// TIA Portal project "DistributoreCaffè" (V19)

(* hardware
DEVICE "S7-1200 station_1"  S7-1200 Station
   slot 0: "Telaio di montaggio_0"  S7-1200 Rack  Rack  V1.0
   slot 1: "PLC"  CPU 1212C DC/DC/Rly  6ES7 212-1HE40-0XB0  V4.6
DEVICE "HMI"  KTP900 Basic PN
   slot 0: "HMI_1"  KTP900 Basic PN  6AV2 123-2JB03-0AX0  17.0.0.0
   slot 1: "HMI_RT_1"  KTP900 Basic PN  6AV2 123-2JB03-0AX0  17.0.0.0
   slot 5: "HMI_1.IE_CP_1"  PROFINET Interface  17.0.0.0
      slot 1: "Interfaccia_1 PROFINET"  PROFINET Interface
         slot 1: "Porta_1"  Port
*)

// ===== PLC "PLC"  CPU 1212C DC/DC/Rly =====

TYPE "CreditoResto"
   STRUCT
      "5Cents" : Real;
      "10Cents" : Real;
      "20Cents" : Real;
      "50Cents" : Real;
      "1Euro" : Real;
      "2Euro" : Real;
   END_STRUCT;
END_TYPE

TYPE "RestoUtente"
   STRUCT
      "5Cents" : SInt;
      "10Cents" : SInt;
      "20Cents" : SInt;
      "50Cents" : SInt;
      "1Euro" : SInt;
      "2Euro" : SInt;
   END_STRUCT;
END_TYPE

TYPE "Prezzo"
   STRUCT
      Bevanda : String;
      Prezzo : Real;
   END_STRUCT;
END_TYPE

DATA_BLOCK "HMI"   // DB1
{ S7_Optimized_Access := 'TRUE' }
VERSION : 0.1
   VAR
      I5cents : Bool;
      I10Cents : Bool;
      I20Cents : Bool;
      I50Cents : Bool;
      I1Euro : Bool;
      I2Euro : Bool;
   END_VAR
   VAR RETAIN
      Resto : "RestoUtente";
   END_VAR
   VAR
      ValvolaBicchiere : Bool;
      ValvolaPaletta : Bool;
      ValvolaCaffè : Bool;
      ValvolaLatte : Bool;
      ValvolaGrappa : Bool;
      ValvolaZucchero : Bool;
      PrelievoProdotto : Bool;
   END_VAR
   VAR RETAIN
      ProdottoPronto : Bool;
   END_VAR
   VAR
      Corto : Bool;
      CortoMacchiato : Bool;
      CortoCorretto : Bool;
      CortoMacchiatoCorretto : Bool;
      Lungo : Bool;
      LungoMacchiato : Bool;
      LungoCorretto : Bool;
      LungoMacchiatoCorretto : Bool;
      ConfermaOrdine : Bool;
      BicchieriScarico : Bool;
      PaletteScarico : Bool;
      CaffèScarico : Bool;
      LatteScarico : Bool;
      GrappaScarico : Bool;
      ZuccheroScarico : Bool;
      Bicchieri : Int;
      Palette : Int;
      Caffè : SInt;
      Latte : SInt;
      Grappa : SInt;
      Zucchero : SInt;
   END_VAR
   VAR RETAIN
      Credito : Real;
      Introiti : Real;
   END_VAR
   VAR
      PrelievoIntroiti : Bool;
      CreditoInsufficiente : Bool;
      QuantitàZuccheroSelezionata : SInt;
      RiduzioneZucchero : Bool;
      IncrementoZucchero : Bool;
      ProdottoInPreparazione : Bool;
   END_VAR
BEGIN
END_DATA_BLOCK

DATA_BLOCK "Sistema"   // DB2
{ S7_Optimized_Access := 'TRUE' }
VERSION : 0.1
   VAR RETAIN
      CreditoResto : "CreditoResto";
   END_VAR
   VAR
      PConfermaOrdine : Bool;
      BloccoInterfacciaUtente : Bool;
      NPrelievoProdotto : Bool;
      BevandaSelezionata : SInt;
      PCorto : Bool;
      PCortoMacchiato : Bool;
      PCortoCorretto : Bool;
      PCortoMacchiatoCorretto : Bool;
      PLungo : Bool;
      PLungoMacchiato : Bool;
      PLungoCorretto : Bool;
      PLungoMacchiatoCorretto : Bool;
      PPiùZucchero : Bool;
      PMenoZucchero : Bool;
   END_VAR
   VAR RETAIN
      Prezzi : Array[1..8] of "Prezzo";
   END_VAR
   VAR
      PBloccoInterfacciaUtente : Bool;
      NPrelievoProdotto2 : Bool;
      NPrelievoIntroiti : Bool;
   END_VAR
BEGIN
   CreditoResto."5Cents" := 5.0;
   CreditoResto."10Cents" := 5.0;
   CreditoResto."20Cents" := 5.0;
   CreditoResto."50Cents" := 5.0;
   CreditoResto."1Euro" := 5.0;
   CreditoResto."2Euro" := 5.0;
   Prezzi[1].Bevanda := 'Corto';
   Prezzi[1].Prezzo := 0.3;
   Prezzi[2].Bevanda := 'CortoMacchiato';
   Prezzi[2].Prezzo := 0.4;
   Prezzi[3].Bevanda := 'CortoCorretto';
   Prezzi[3].Prezzo := 0.4;
   Prezzi[4].Bevanda := 'CortoMacchiatoCorretto';
   Prezzi[4].Prezzo := 0.5;
   Prezzi[5].Bevanda := 'Lungo';
   Prezzi[5].Prezzo := 0.6;
   Prezzi[6].Bevanda := 'LungoMacchiato';
   Prezzi[6].Prezzo := 0.7;
   Prezzi[7].Bevanda := 'LungoCorretto';
   Prezzi[7].Prezzo := 0.7;
   Prezzi[8].Bevanda := 'LungoMacchiatoCorretto';
   Prezzi[8].Prezzo := 0.8;
END_DATA_BLOCK

DATA_BLOCK "AggiornamentoCreditoUtente_DB"   // DB3
{ S7_Optimized_Access := 'TRUE' }
VERSION : 0.1
// stored: InstanceOfName AggiornamentoCreditoUtenteCreditoDistributore
"AggiornamentoCreditoUtenteCreditoDistributore"
BEGIN
END_DATA_BLOCK

DATA_BLOCK "PreparazioneBevanda_DB"   // DB4
{ S7_Optimized_Access := 'TRUE' }
VERSION : 0.1
// stored: InstanceOfName PreparazioneBevanda
"PreparazioneBevanda"
BEGIN
END_DATA_BLOCK

DATA_BLOCK "AggiornamentoRestoUtenteCreditoUtenteCreditoDistributore_DB"   // DB5
{ S7_Optimized_Access := 'TRUE' }
VERSION : 0.1
// stored: InstanceOfName AggiornamentoRestoUtenteCreditoUtenteCreditoDistributore
"AggiornamentoRestoUtenteCreditoUtenteCreditoDistributore"
BEGIN
END_DATA_BLOCK

FUNCTION_BLOCK "AggiornamentoCreditoUtenteCreditoDistributore"   // FB1, LAD
{ S7_Optimized_Access := 'TRUE' }
VERSION : 0.1
   VAR_INPUT
      "5Cents" : Bool;
      "10Cents" : Bool;
      "20Cents" : Bool;
      "50Cents" : Bool;
      "1Euro" : Bool;
      "2Euro" : Bool;
   END_VAR
   VAR_IN_OUT
      CreditoDistributore : "CreditoResto";
      CreditoUtente : Real;
   END_VAR
   VAR
      PI5Cents : Bool;
      PI10Cents : Bool;
      PI20Cents : Bool;
      PI50Cents : Bool;
      PI1Euro : Bool;
      PI2Euro : Bool;
   END_VAR
   VAR_TEMP   // added for the SCL form of the ladder/FBD networks
      _w1 : Bool;
      _w2 : Bool;
      _w3 : Bool;
      _w4 : Bool;
      _w5 : Bool;
      _w6 : Bool;
   END_VAR
BEGIN

REGION Network 1
   // Attenzione: i valori Real non sempre vengono salvati a cifra tonda
   // (Es: 0.2999999999.. oppure 0.31111111.. invece di 0.3)
   // Arrotondare dopo ogni operazione matematica che li implica
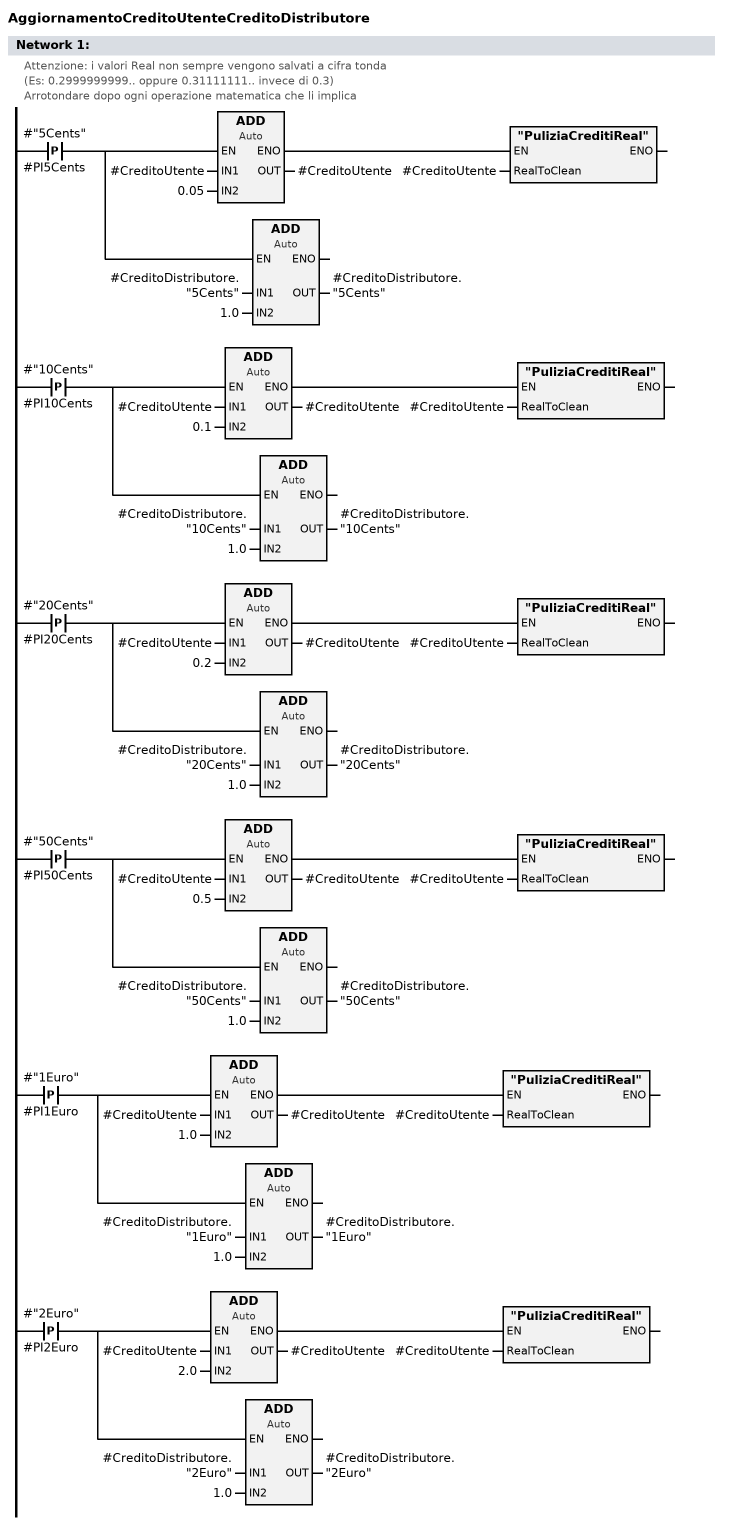
   RUNG wire#powerrail
      P_Contact(operand := #"5Cents", bit := #PI5Cents)
      wire#w1
      Add(in1 := #CreditoUtente, in2 := 0.05, out => #CreditoUtente)
      "PuliziaCreditiReal"(RealToClean := #CreditoUtente)
   END_RUNG
   RUNG wire#w1
      Add(in1 := #CreditoDistributore."5Cents", in2 := 1.0, out => #CreditoDistributore."5Cents")
   END_RUNG
   RUNG wire#powerrail
      P_Contact(operand := #"10Cents", bit := #PI10Cents)
      wire#w2
      Add(in1 := #CreditoUtente, in2 := 0.1, out => #CreditoUtente)
      "PuliziaCreditiReal"(RealToClean := #CreditoUtente)
   END_RUNG
   RUNG wire#w2
      Add(in1 := #CreditoDistributore."10Cents", in2 := 1.0, out => #CreditoDistributore."10Cents")
   END_RUNG
   RUNG wire#powerrail
      P_Contact(operand := #"20Cents", bit := #PI20Cents)
      wire#w3
      Add(in1 := #CreditoUtente, in2 := 0.2, out => #CreditoUtente)
      "PuliziaCreditiReal"(RealToClean := #CreditoUtente)
   END_RUNG
   RUNG wire#w3
      Add(in1 := #CreditoDistributore."20Cents", in2 := 1.0, out => #CreditoDistributore."20Cents")
   END_RUNG
   RUNG wire#powerrail
      P_Contact(operand := #"50Cents", bit := #PI50Cents)
      wire#w4
      Add(in1 := #CreditoUtente, in2 := 0.5, out => #CreditoUtente)
      "PuliziaCreditiReal"(RealToClean := #CreditoUtente)
   END_RUNG
   RUNG wire#w4
      Add(in1 := #CreditoDistributore."50Cents", in2 := 1.0, out => #CreditoDistributore."50Cents")
   END_RUNG
   RUNG wire#powerrail
      P_Contact(operand := #"1Euro", bit := #PI1Euro)
      wire#w5
      Add(in1 := #CreditoUtente, in2 := 1.0, out => #CreditoUtente)
      "PuliziaCreditiReal"(RealToClean := #CreditoUtente)
   END_RUNG
   RUNG wire#w5
      Add(in1 := #CreditoDistributore."1Euro", in2 := 1.0, out => #CreditoDistributore."1Euro")
   END_RUNG
   RUNG wire#powerrail
      P_Contact(operand := #"2Euro", bit := #PI2Euro)
      wire#w6
      Add(in1 := #CreditoUtente, in2 := 2.0, out => #CreditoUtente)
      "PuliziaCreditiReal"(RealToClean := #CreditoUtente)
   END_RUNG
   RUNG wire#w6
      Add(in1 := #CreditoDistributore."2Euro", in2 := 1.0, out => #CreditoDistributore."2Euro")
   END_RUNG
   // the same network as SCL:
   #_w1 := #"5Cents" AND NOT #PI5Cents;   // rising edge of #"5Cents"
   #PI5Cents := #"5Cents";
   IF #_w1 THEN
       #CreditoUtente := #CreditoUtente + 0.05;
       "PuliziaCreditiReal"(RealToClean := #CreditoUtente);
       #CreditoDistributore."5Cents" := #CreditoDistributore."5Cents" + 1.0;
   END_IF;
   #_w2 := #"10Cents" AND NOT #PI10Cents;   // rising edge of #"10Cents"
   #PI10Cents := #"10Cents";
   IF #_w2 THEN
       #CreditoUtente := #CreditoUtente + 0.1;
       "PuliziaCreditiReal"(RealToClean := #CreditoUtente);
       #CreditoDistributore."10Cents" := #CreditoDistributore."10Cents" + 1.0;
   END_IF;
   #_w3 := #"20Cents" AND NOT #PI20Cents;   // rising edge of #"20Cents"
   #PI20Cents := #"20Cents";
   IF #_w3 THEN
       #CreditoUtente := #CreditoUtente + 0.2;
       "PuliziaCreditiReal"(RealToClean := #CreditoUtente);
       #CreditoDistributore."20Cents" := #CreditoDistributore."20Cents" + 1.0;
   END_IF;
   #_w4 := #"50Cents" AND NOT #PI50Cents;   // rising edge of #"50Cents"
   #PI50Cents := #"50Cents";
   IF #_w4 THEN
       #CreditoUtente := #CreditoUtente + 0.5;
       "PuliziaCreditiReal"(RealToClean := #CreditoUtente);
       #CreditoDistributore."50Cents" := #CreditoDistributore."50Cents" + 1.0;
   END_IF;
   #_w5 := #"1Euro" AND NOT #PI1Euro;   // rising edge of #"1Euro"
   #PI1Euro := #"1Euro";
   IF #_w5 THEN
       #CreditoUtente := #CreditoUtente + 1.0;
       "PuliziaCreditiReal"(RealToClean := #CreditoUtente);
       #CreditoDistributore."1Euro" := #CreditoDistributore."1Euro" + 1.0;
   END_IF;
   #_w6 := #"2Euro" AND NOT #PI2Euro;   // rising edge of #"2Euro"
   #PI2Euro := #"2Euro";
   IF #_w6 THEN
       #CreditoUtente := #CreditoUtente + 2.0;
       "PuliziaCreditiReal"(RealToClean := #CreditoUtente);
       #CreditoDistributore."2Euro" := #CreditoDistributore."2Euro" + 1.0;
   END_IF;
END_REGION
END_FUNCTION_BLOCK

FUNCTION_BLOCK "PreparazioneBevanda"   // FB2, LAD
{ S7_Optimized_Access := 'TRUE' }
VERSION : 0.1
   VAR_INPUT
      BevandaSelezionata : SInt;
      InnescoProcesso : Bool;
   END_VAR
   VAR
      TPBicchiere : TP_TIME;
      NQTPBicchiere : Bool;
      TPPaletta : TP_TIME;
      NQTPPaletta : Bool;
      TPCaffè : TP_TIME;
      NQTPCaffè : Bool;
      TPLatte : TP_TIME;
      NQTPLatte : Bool;
      TPGrappa : TP_TIME;
      NQTPGrappa : Bool;
      TPzucchero : TP_TIME;
      NQTPZucchero : Bool;
      PInnescoProcesso : Bool;
   END_VAR
   VAR_TEMP
      PTZucchero : Int;
   END_VAR
   VAR_TEMP   // added for the SCL form of the ladder/FBD networks
      _w1 : Bool;
      _w2 : Bool;
      _w3 : Bool;
      _w4 : Bool;
      _w5 : Bool;
      _w6 : Bool;
      _w7 : Bool;
      _w8 : Bool;
      _w9 : Bool;
      _w10 : Bool;
      _w11 : Bool;
      _w12 : Bool;
   END_VAR
BEGIN

REGION Network 1
   // Gestire trigger timer valvole
   // - grappa caso bevanda corretta non macchiata
   // - zucchero caso bevanda zuccherata liscia o macchiata
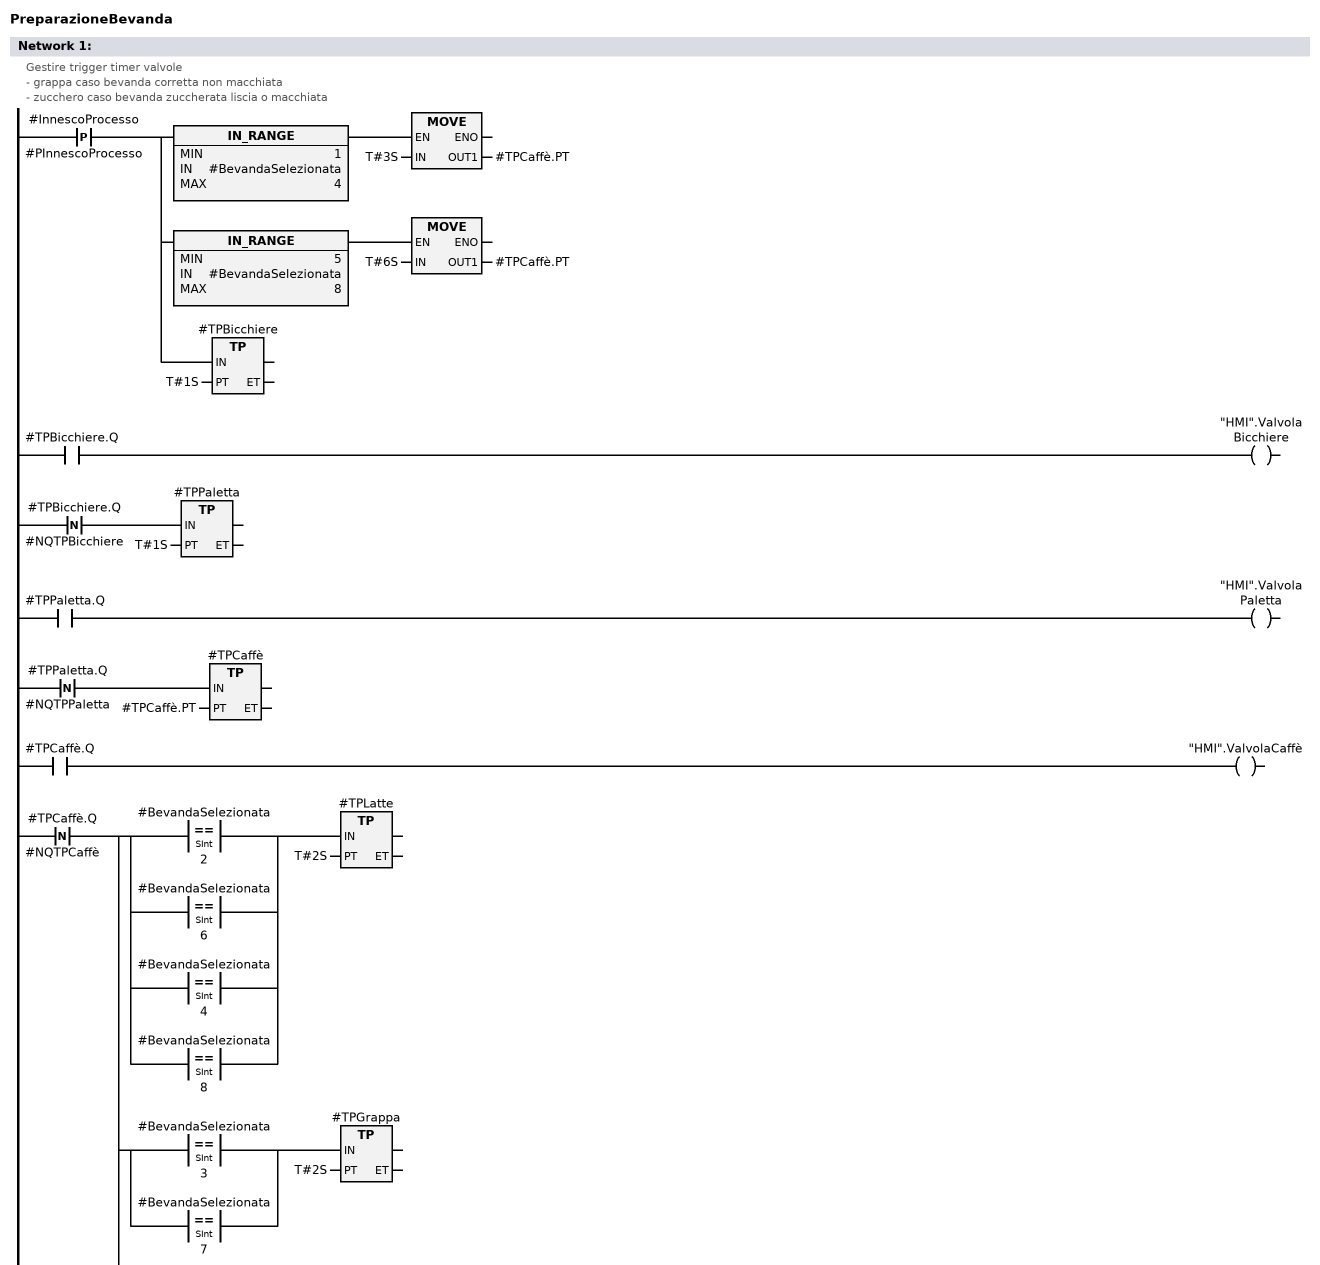
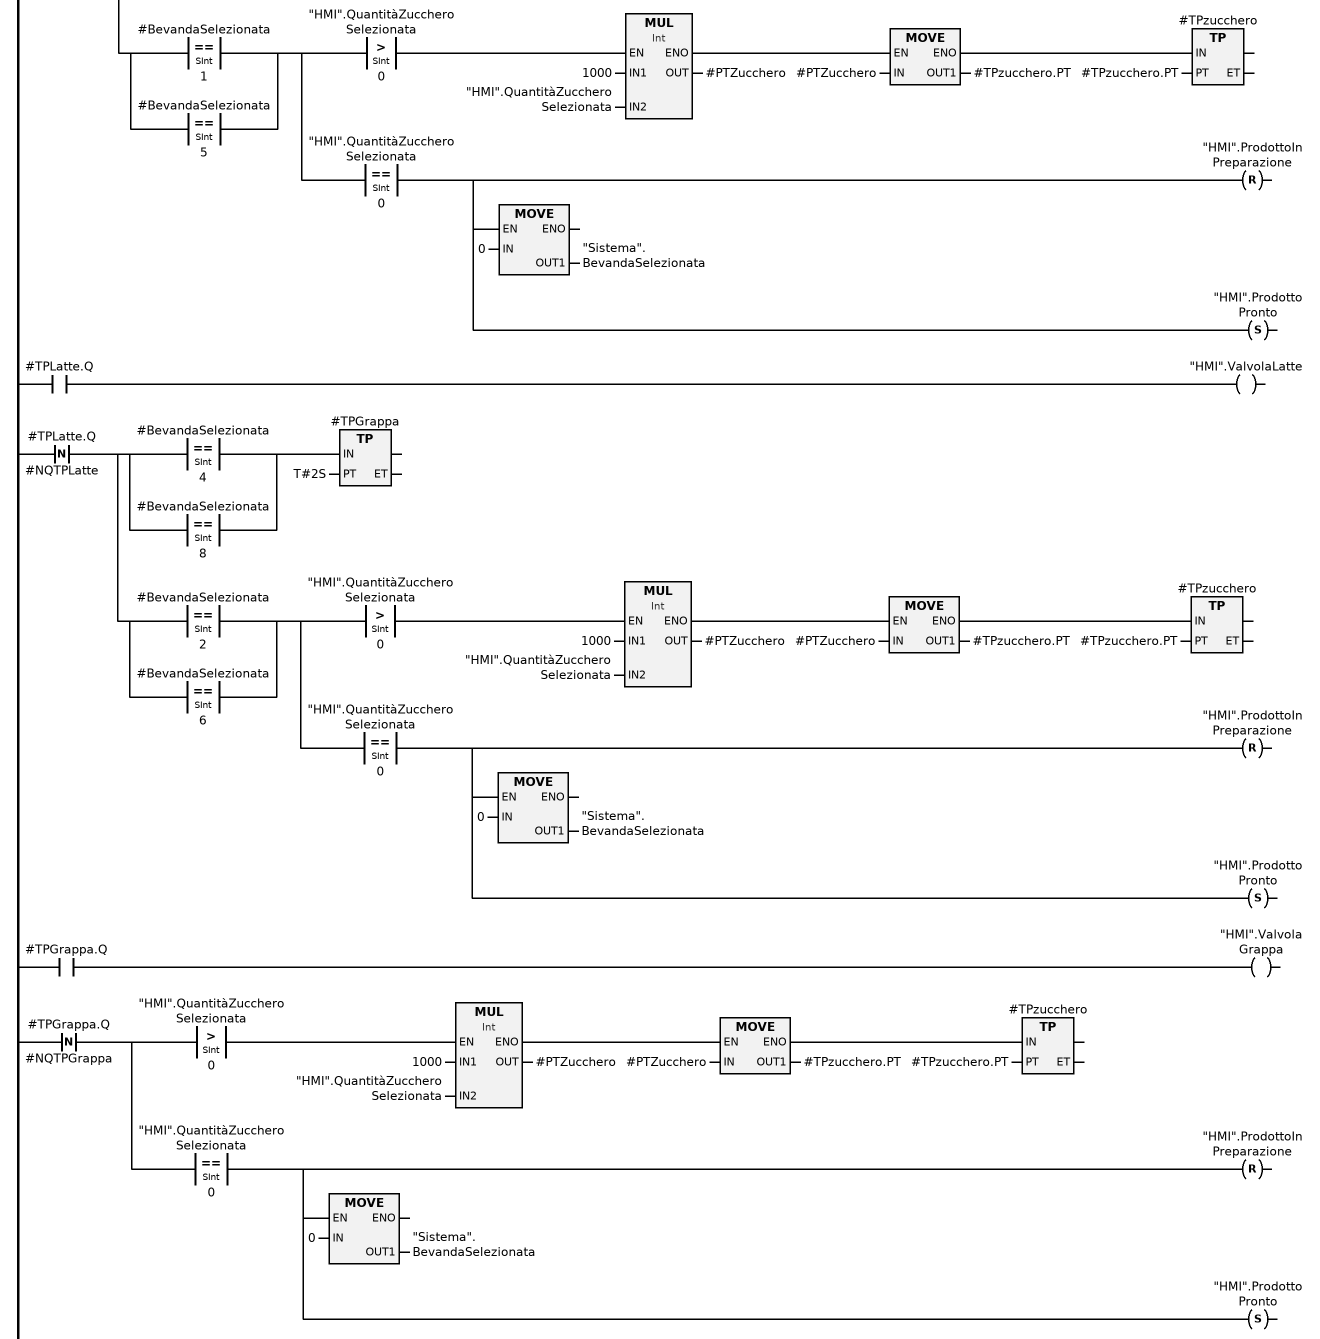
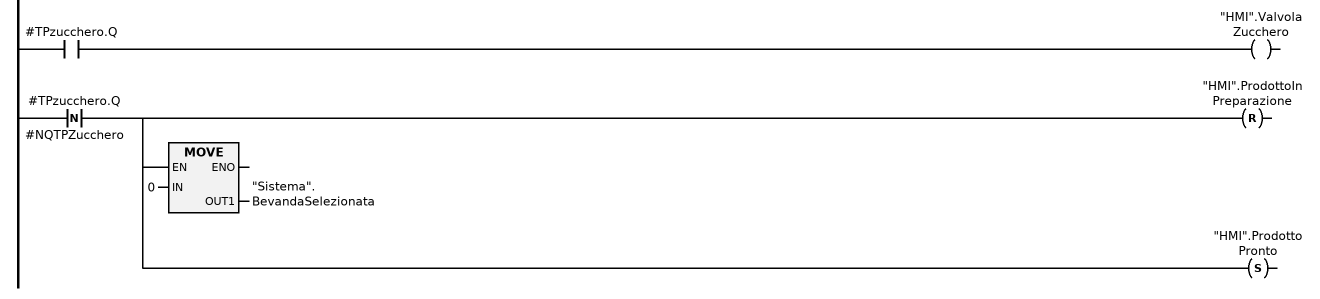
   #_w1 := #InnescoProcesso AND NOT #PInnescoProcesso;   // rising edge of #InnescoProcesso
   #PInnescoProcesso := #InnescoProcesso;
   IF #_w1 AND (1 <= #BevandaSelezionata) AND (#BevandaSelezionata <= 4) THEN #TPCaffè.PT := T#3S; END_IF;
   IF #_w1 AND (5 <= #BevandaSelezionata) AND (#BevandaSelezionata <= 8) THEN #TPCaffè.PT := T#6S; END_IF;
   #TPBicchiere(IN := #_w1, PT := T#1S);   // TP
   "HMI".ValvolaBicchiere := #TPBicchiere.Q;
   #_w2 := NOT #TPBicchiere.Q AND #NQTPBicchiere;   // falling edge of #TPBicchiere.Q
   #NQTPBicchiere := #TPBicchiere.Q;
   #TPPaletta(IN := #_w2, PT := T#1S);   // TP
   "HMI".ValvolaPaletta := #TPPaletta.Q;
   #_w3 := NOT #TPPaletta.Q AND #NQTPPaletta;   // falling edge of #TPPaletta.Q
   #NQTPPaletta := #TPPaletta.Q;
   #TPCaffè(IN := #_w3, PT := #TPCaffè.PT);   // TP
   "HMI".ValvolaCaffè := #TPCaffè.Q;
   #_w4 := NOT #TPCaffè.Q AND #NQTPCaffè;   // falling edge of #TPCaffè.Q
   #NQTPCaffè := #TPCaffè.Q;
   #TPLatte(IN := #_w4 AND ((#BevandaSelezionata = 2) OR (#BevandaSelezionata = 6) OR (#BevandaSelezionata = 4) OR (#BevandaSelezionata = 8)),   // TP
            PT := T#2S);
   #TPGrappa(IN := #_w4 AND ((#BevandaSelezionata = 3) OR (#BevandaSelezionata = 7)), PT := T#2S);   // TP
   #_w5 := #_w4 AND ((#BevandaSelezionata = 1) OR (#BevandaSelezionata = 5));
   #_w6 := #_w5 AND ("HMI".QuantitàZuccheroSelezionata > 0);
   IF #_w6 THEN
       #PTZucchero := 1000 * "HMI".QuantitàZuccheroSelezionata;
       #TPzucchero.PT := #PTZucchero;
   END_IF;
   #TPzucchero(IN := #_w6, PT := #TPzucchero.PT);   // TP
   IF #_w5 AND ("HMI".QuantitàZuccheroSelezionata = 0) THEN
       "HMI".ProdottoInPreparazione := FALSE;
       "Sistema".BevandaSelezionata := 0;
       "HMI".ProdottoPronto := TRUE;
   END_IF;
   "HMI".ValvolaLatte := #TPLatte.Q;
   #_w7 := NOT #TPLatte.Q AND #NQTPLatte;   // falling edge of #TPLatte.Q
   #NQTPLatte := #TPLatte.Q;
   #TPGrappa(IN := #_w7 AND ((#BevandaSelezionata = 4) OR (#BevandaSelezionata = 8)), PT := T#2S);   // TP
   #_w8 := #_w7 AND ((#BevandaSelezionata = 2) OR (#BevandaSelezionata = 6));
   #_w9 := #_w8 AND ("HMI".QuantitàZuccheroSelezionata > 0);
   IF #_w9 THEN
       #PTZucchero := 1000 * "HMI".QuantitàZuccheroSelezionata;
       #TPzucchero.PT := #PTZucchero;
   END_IF;
   #TPzucchero(IN := #_w9, PT := #TPzucchero.PT);   // TP
   IF #_w8 AND ("HMI".QuantitàZuccheroSelezionata = 0) THEN
       "HMI".ProdottoInPreparazione := FALSE;
       "Sistema".BevandaSelezionata := 0;
       "HMI".ProdottoPronto := TRUE;
   END_IF;
   "HMI".ValvolaGrappa := #TPGrappa.Q;
   #_w10 := NOT #TPGrappa.Q AND #NQTPGrappa;   // falling edge of #TPGrappa.Q
   #NQTPGrappa := #TPGrappa.Q;
   #_w11 := #_w10 AND ("HMI".QuantitàZuccheroSelezionata > 0);
   IF #_w11 THEN
       #PTZucchero := 1000 * "HMI".QuantitàZuccheroSelezionata;
       #TPzucchero.PT := #PTZucchero;
   END_IF;
   #TPzucchero(IN := #_w11, PT := #TPzucchero.PT);   // TP
   IF #_w10 AND ("HMI".QuantitàZuccheroSelezionata = 0) THEN
       "HMI".ProdottoInPreparazione := FALSE;
       "Sistema".BevandaSelezionata := 0;
       "HMI".ProdottoPronto := TRUE;
   END_IF;
   "HMI".ValvolaZucchero := #TPzucchero.Q;
   #_w12 := NOT #TPzucchero.Q AND #NQTPZucchero;   // falling edge of #TPzucchero.Q
   #NQTPZucchero := #TPzucchero.Q;
   IF #_w12 THEN
       "HMI".ProdottoInPreparazione := FALSE;
       "Sistema".BevandaSelezionata := 0;
       "HMI".ProdottoPronto := TRUE;
   END_IF;
END_REGION
END_FUNCTION_BLOCK

FUNCTION_BLOCK "AggiornamentoRestoUtenteCreditoUtenteCreditoDistributore"   // FB3, SCL
{ S7_Optimized_Access := 'TRUE' }
VERSION : 0.1
   VAR_INPUT
      BevandaSelezionata : SInt;
      InnescoProcesso : Bool;
   END_VAR
   VAR_IN_OUT
      Resto : "RestoUtente";
      CreditoDistributore : "CreditoResto";
      CreditoUtente : Real;
   END_VAR
   VAR
      Inception_R_TRIG_Instance : R_TRIG;
   END_VAR
BEGIN
   #Inception_R_TRIG_Instance(CLK:=#InnescoProcesso,
                              Q=>#Inception_R_TRIG_Instance.Q);

   IF #Inception_R_TRIG_Instance.Q THEN
       // Attenzione: i valori Real non sempre vengono salvati a cifra tonda
       // (Es: 0.2999999999.. oppure 0.31111111.. invece di 0.3)
       // Arrotondare dopo ogni operazione matematica che li implica
       #CreditoUtente := #CreditoUtente - "Sistema".Prezzi[#BevandaSelezionata].Prezzo;
       #CreditoUtente := DINT_TO_REAL(ROUND(#CreditoUtente * 100.0)) / 100.0;

       // Quantizzazione resto nei tagli di moneta disponibili nel salvadanaio del distributore
       // fino ad azzeramento credito utente residuo
       // Qualora il credito distributore sia insufficiente il credito utente residuo resta disponibile
       // per i prossimi acquisti
       WHILE #CreditoUtente >= 2.0 DO
           IF #CreditoDistributore."2Euro" > 0 THEN // (I tipi di monete inseriti dall'utenza sono già confluiti nel credito del distributore)
               // Rimuovere monete dal credito distributore...
               #CreditoDistributore."2Euro" := #CreditoDistributore."2Euro" - 1.0;
               // ... Aggiungerle al resto utente
               #Resto."2Euro" := #Resto."2Euro" + 1;
               // Aggiornare credito utente residuo
               #CreditoUtente := #CreditoUtente - 2.0;
               "PuliziaCreditiReal"(#CreditoUtente);
           ELSIF #CreditoDistributore."1Euro" > 0 THEN
               // Rimuovere monete dal credito distributore...
               #CreditoDistributore."1Euro" := #CreditoDistributore."1Euro" - 1.0;
               // ... Aggiungerle al resto utente
               #Resto."1Euro" := #Resto."1Euro" + 1;
               // Aggiornare credito utente residuo
               #CreditoUtente := #CreditoUtente - 1.0;
               "PuliziaCreditiReal"(#CreditoUtente);
           ELSIF #CreditoDistributore."50Cents" > 0 THEN
               #CreditoDistributore."50Cents" := #CreditoDistributore."50Cents" - 1.0;
               #Resto."50Cents" := #Resto."50Cents" + 1;
               #CreditoUtente := #CreditoUtente - 0.5;
               "PuliziaCreditiReal"(#CreditoUtente);
           ELSIF #CreditoDistributore."20Cents" > 0 THEN
               #CreditoDistributore."20Cents" := #CreditoDistributore."20Cents" - 1.0;
               #Resto."20Cents" := #Resto."20Cents" + 1;
               #CreditoUtente := #CreditoUtente - 0.2;
               "PuliziaCreditiReal"(#CreditoUtente);
           ELSIF #CreditoDistributore."10Cents" > 0 THEN
               #CreditoDistributore."10Cents" := #CreditoDistributore."10Cents" - 1.0;
               #Resto."10Cents" := #Resto."10Cents" + 1;
               #CreditoUtente := #CreditoUtente - 0.1;
               "PuliziaCreditiReal"(#CreditoUtente);
           ELSIF #CreditoDistributore."5Cents" > 0 THEN
               #CreditoDistributore."5Cents" := #CreditoDistributore."5Cents" - 1.0;
               #Resto."5Cents" := #Resto."5Cents" + 1;
               #CreditoUtente := #CreditoUtente - 0.05;
               "PuliziaCreditiReal"(#CreditoUtente);
           END_IF;
       END_WHILE;

       WHILE #CreditoUtente >= 1.0 DO
           IF #CreditoDistributore."1Euro" > 0 THEN
               #CreditoDistributore."1Euro" := #CreditoDistributore."1Euro" - 1.0;
               #Resto."1Euro" := #Resto."1Euro" + 1;
               #CreditoUtente := #CreditoUtente - 1.0;
               "PuliziaCreditiReal"(#CreditoUtente);
           ELSIF #CreditoDistributore."50Cents" > 0 THEN
               #CreditoDistributore."50Cents" := #CreditoDistributore."50Cents" - 1.0;
               #Resto."50Cents" := #Resto."50Cents" + 1;
               #CreditoUtente := #CreditoUtente - 0.5;
               "PuliziaCreditiReal"(#CreditoUtente);
           ELSIF #CreditoDistributore."20Cents" > 0 THEN
               #CreditoDistributore."20Cents" := #CreditoDistributore."20Cents" - 1.0;
               #Resto."20Cents" := #Resto."20Cents" + 1;
               #CreditoUtente := #CreditoUtente - 0.2;
               "PuliziaCreditiReal"(#CreditoUtente);
           ELSIF #CreditoDistributore."10Cents" > 0 THEN
               #CreditoDistributore."10Cents" := #CreditoDistributore."10Cents" - 1.0;
               #Resto."10Cents" := #Resto."10Cents" + 1;
               #CreditoUtente := #CreditoUtente - 0.1;
               "PuliziaCreditiReal"(#CreditoUtente);
           ELSIF #CreditoDistributore."5Cents" > 0 THEN
               #CreditoDistributore."5Cents" := #CreditoDistributore."5Cents" - 1.0;
               #Resto."5Cents" := #Resto."5Cents" + 1;
               #CreditoUtente := #CreditoUtente - 0.05;
               "PuliziaCreditiReal"(#CreditoUtente);
           END_IF;
       END_WHILE;

       WHILE #CreditoUtente >= 0.5 DO
           IF #CreditoDistributore."50Cents" > 0 THEN
               #CreditoDistributore."50Cents" := #CreditoDistributore."50Cents" - 1.0;
               #Resto."50Cents" := #Resto."50Cents" + 1;
               #CreditoUtente := #CreditoUtente - 0.5;
               "PuliziaCreditiReal"(#CreditoUtente);
           ELSIF #CreditoDistributore."20Cents" > 0 THEN
               #CreditoDistributore."20Cents" := #CreditoDistributore."20Cents" - 1.0;
               #Resto."20Cents" := #Resto."20Cents" + 1;
               #CreditoUtente := #CreditoUtente - 0.2;
               "PuliziaCreditiReal"(#CreditoUtente);
           ELSIF #CreditoDistributore."10Cents" > 0 THEN
               #CreditoDistributore."10Cents" := #CreditoDistributore."10Cents" - 1.0;
               #Resto."10Cents" := #Resto."10Cents" + 1;
               #CreditoUtente := #CreditoUtente - 0.1;
               "PuliziaCreditiReal"(#CreditoUtente);
           ELSIF #CreditoDistributore."5Cents" > 0 THEN
               #CreditoDistributore."5Cents" := #CreditoDistributore."5Cents" - 1.0;
               #Resto."5Cents" := #Resto."5Cents" + 1;
               #CreditoUtente := #CreditoUtente - 0.05;
               "PuliziaCreditiReal"(#CreditoUtente);
           END_IF;
       END_WHILE;

       WHILE #CreditoUtente >= 0.2 DO
           IF #CreditoDistributore."20Cents" > 0 THEN
               #CreditoDistributore."20Cents" := #CreditoDistributore."20Cents" - 1.0;
               #Resto."20Cents" := #Resto."20Cents" + 1;
               #CreditoUtente := #CreditoUtente - 0.2;
               "PuliziaCreditiReal"(#CreditoUtente);
           ELSIF #CreditoDistributore."10Cents" > 0 THEN
               #CreditoDistributore."10Cents" := #CreditoDistributore."10Cents" - 1.0;
               #Resto."10Cents" := #Resto."10Cents" + 1;
               #CreditoUtente := #CreditoUtente - 0.1;
               "PuliziaCreditiReal"(#CreditoUtente);
           ELSIF #CreditoDistributore."5Cents" > 0 THEN
               #CreditoDistributore."5Cents" := #CreditoDistributore."5Cents" - 1.0;
               #Resto."5Cents" := #Resto."5Cents" + 1;
               #CreditoUtente := #CreditoUtente - 0.05;
               "PuliziaCreditiReal"(#CreditoUtente);
           END_IF;
       END_WHILE;

       WHILE #CreditoUtente >= 0.1 DO
           IF #CreditoDistributore."10Cents" > 0 THEN
               #CreditoDistributore."10Cents" := #CreditoDistributore."10Cents" - 1.0;
               #Resto."10Cents" := #Resto."10Cents" + 1;
               #CreditoUtente := #CreditoUtente - 0.1;
               "PuliziaCreditiReal"(#CreditoUtente);
           ELSIF #CreditoDistributore."5Cents" > 0 THEN
               #CreditoDistributore."5Cents" := #CreditoDistributore."5Cents" - 1.0;
               #Resto."5Cents" := #Resto."5Cents" + 1;
               #CreditoUtente := #CreditoUtente - 0.05;
               "PuliziaCreditiReal"(#CreditoUtente);
           END_IF;
       END_WHILE;

       WHILE #CreditoUtente >= 0.05 DO
           IF #CreditoDistributore."5Cents" > 0 THEN
               #CreditoDistributore."5Cents" := #CreditoDistributore."5Cents" - 1.0;
               #Resto."5Cents" := #Resto."5Cents" + 1;
               #CreditoUtente := #CreditoUtente - 0.05;
               "PuliziaCreditiReal"(#CreditoUtente);
           END_IF;
       END_WHILE;

       // Aggiornamento introiti proprietario
       "AggiornamentoIntroiti"(CreditoDistributore:="Sistema".CreditoResto,
                               Introiti:="HMI".Introiti);

   END_IF;
END_FUNCTION_BLOCK

FUNCTION "AggiornamentoIntroiti" : Void   // FC1, SCL
{ S7_Optimized_Access := 'TRUE' }
VERSION : 0.1
   VAR_INPUT
      CreditoDistributore : "CreditoResto";
   END_VAR
   VAR_IN_OUT
      Introiti : Real;
   END_VAR
   VAR CONSTANT
      CreditoIniziale : Real := 19.25;
   END_VAR
BEGIN
   // Il credito iniziale, destinato all'erogazione agevolata del resto, non costituisce guadagno per il proprietario

   // Attenzione: i valori Real non sempre vengono salvati a cifra tonda
   // (Es: 0.2999999999.. oppure 0.31111111.. invece di 0.3)
   // Arrotondare dopo ogni operazione matematica che li implica

   #Introiti := #CreditoDistributore."2Euro" * 2.0 + #CreditoDistributore."1Euro" + #CreditoDistributore."50Cents" * 0.5 + #CreditoDistributore."20Cents" * 0.2 + #CreditoDistributore."10Cents" * 0.1 + #CreditoDistributore."5Cents" * 0.05 - #CreditoIniziale;
   "PuliziaCreditiReal"(#Introiti);
END_FUNCTION

FUNCTION "ValutazioneInsufficienzaCredito" : Void   // FC2, SCL
{ S7_Optimized_Access := 'TRUE' }
VERSION : 0.1
   VAR_INPUT
      BevandaSelezionata : SInt;
      CreditoUtente : Real;
   END_VAR
   VAR_IN_OUT
      CreditoInsufficiente : Bool;
   END_VAR
BEGIN
   IF #CreditoUtente < ("Sistema".Prezzi[#BevandaSelezionata].Prezzo) THEN
       #CreditoInsufficiente := TRUE;
   ELSE
       #CreditoInsufficiente := FALSE;
   END_IF;
END_FUNCTION

FUNCTION "PuliziaCreditiReal" : Void   // FC3, SCL
{ S7_Optimized_Access := 'TRUE' }
VERSION : 0.1
   VAR_IN_OUT
      RealToClean : Real;
   END_VAR
BEGIN
   #RealToClean := DINT_TO_REAL(ROUND(#RealToClean * 100.0)) / 100.0; // (ROUND() restituisce D/INT)
   // (moltiplicazione/divisione per potenze di 10 non dovrebbe dare origine a decimali sporchi)
END_FUNCTION

ORGANIZATION_BLOCK "Main"   // OB1, LAD, ProgramCycle
TITLE = "Main Program Sweep (Cycle)"
{ S7_Optimized_Access := 'TRUE' }
VERSION : 0.1
   VAR_INPUT
      Initial_Call : Bool;   // Initial call of this OB
      Remanence : Bool;   // =True, if remanent data are available
   END_VAR
   VAR_TEMP   // added for the SCL form of the ladder/FBD networks
      _w1 : Bool;
      _w2 : Bool;
      _w3 : Bool;
      _w4 : Bool;
      _w5 : Bool;
      _w6 : Bool;
      _w7 : Bool;
      _w8 : Bool;
      _w9 : Bool;
   END_VAR
BEGIN

REGION Network 1
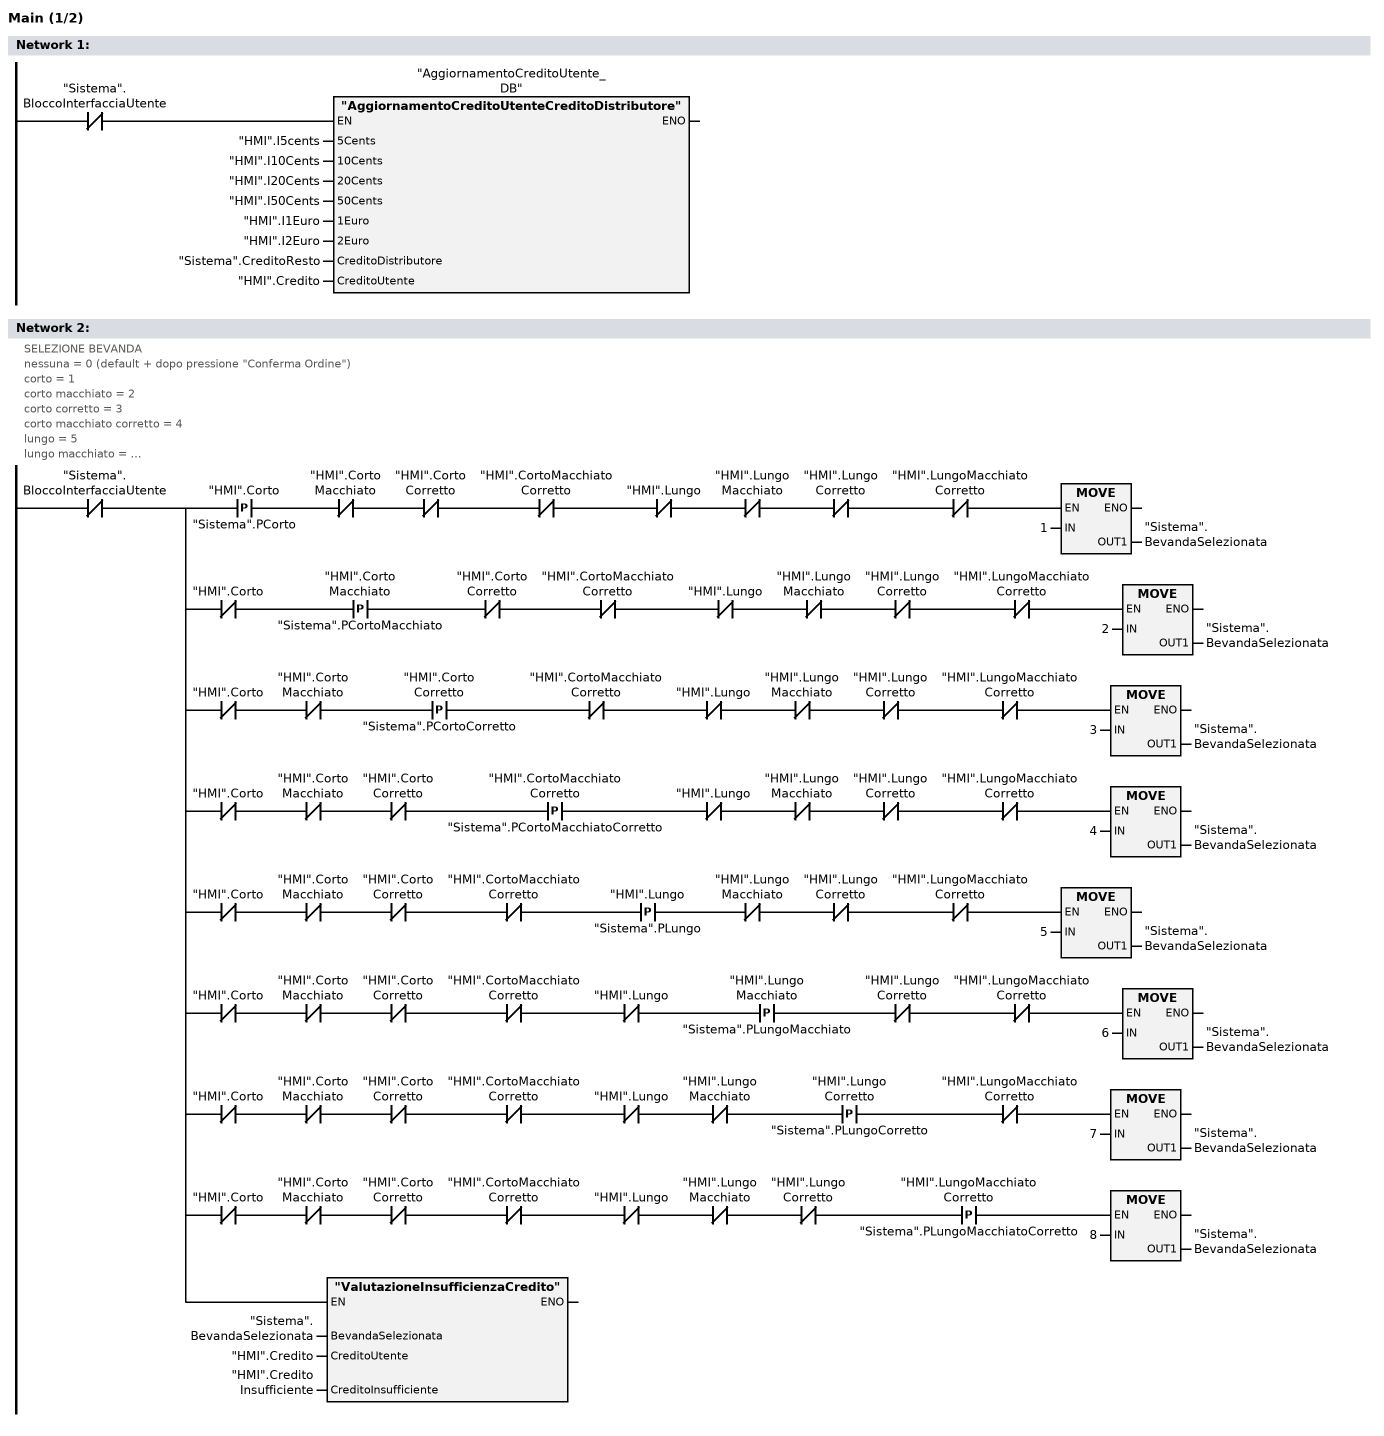
   RUNG wire#powerrail
      I_Contact( "Sistema".BloccoInterfacciaUtente )
      "AggiornamentoCreditoUtente_DB"("5Cents" := "HMI".I5cents, "10Cents" := "HMI".I10Cents, "20Cents" := "HMI".I20Cents, "50Cents" := "HMI".I50Cents, "1Euro" := "HMI".I1Euro, "2Euro" := "HMI".I2Euro, CreditoDistributore := "Sistema".CreditoResto, CreditoUtente := "HMI".Credito)
   END_RUNG
   // the same network as SCL:
   IF NOT "Sistema".BloccoInterfacciaUtente THEN
       "AggiornamentoCreditoUtente_DB"("5Cents" := "HMI".I5cents,   // "AggiornamentoCreditoUtenteCreditoDistributore"
                               "10Cents" := "HMI".I10Cents,
                               "20Cents" := "HMI".I20Cents,
                               "50Cents" := "HMI".I50Cents,
                               "1Euro" := "HMI".I1Euro,
                               "2Euro" := "HMI".I2Euro,
                               CreditoDistributore := "Sistema".CreditoResto,
                               CreditoUtente := "HMI".Credito);
   END_IF;
END_REGION

REGION Network 2
   // SELEZIONE BEVANDA
   // 
   // nessuna = 0 (default + dopo pressione "Conferma Ordine")
   // corto = 1
   // corto macchiato = 2
   // corto corretto = 3
   // corto macchiato corretto = 4
   // lungo = 5
   // lungo macchiato = 6
   // lungo corretto = 7
   // lungo macchiato corretto = 8
   // 
   // Il distributore avvisa con un lampeggio del diplay credito l'insufficienza di credito
   // 
   // Caso più pulsanti premuti contemporaneamente: priorità primo premuto
   RUNG wire#powerrail
      I_Contact( "Sistema".BloccoInterfacciaUtente )
      wire#w1
      P_Contact(operand := "HMI".Corto, bit := "Sistema".PCorto)
      I_Contact( "HMI".CortoMacchiato )
      I_Contact( "HMI".CortoCorretto )
      I_Contact( "HMI".CortoMacchiatoCorretto )
      I_Contact( "HMI".Lungo )
      I_Contact( "HMI".LungoMacchiato )
      I_Contact( "HMI".LungoCorretto )
      I_Contact( "HMI".LungoMacchiatoCorretto )
      Move(in := 1, out1 => "Sistema".BevandaSelezionata)
   END_RUNG
   RUNG wire#w1
      I_Contact( "HMI".Corto )
      P_Contact(operand := "HMI".CortoMacchiato, bit := "Sistema".PCortoMacchiato)
      I_Contact( "HMI".CortoCorretto )
      I_Contact( "HMI".CortoMacchiatoCorretto )
      I_Contact( "HMI".Lungo )
      I_Contact( "HMI".LungoMacchiato )
      I_Contact( "HMI".LungoCorretto )
      I_Contact( "HMI".LungoMacchiatoCorretto )
      Move(in := 2, out1 => "Sistema".BevandaSelezionata)
   END_RUNG
   RUNG wire#w1
      I_Contact( "HMI".Corto )
      I_Contact( "HMI".CortoMacchiato )
      P_Contact(operand := "HMI".CortoCorretto, bit := "Sistema".PCortoCorretto)
      I_Contact( "HMI".CortoMacchiatoCorretto )
      I_Contact( "HMI".Lungo )
      I_Contact( "HMI".LungoMacchiato )
      I_Contact( "HMI".LungoCorretto )
      I_Contact( "HMI".LungoMacchiatoCorretto )
      Move(in := 3, out1 => "Sistema".BevandaSelezionata)
   END_RUNG
   RUNG wire#w1
      I_Contact( "HMI".Corto )
      I_Contact( "HMI".CortoMacchiato )
      I_Contact( "HMI".CortoCorretto )
      P_Contact(operand := "HMI".CortoMacchiatoCorretto, bit := "Sistema".PCortoMacchiatoCorretto)
      I_Contact( "HMI".Lungo )
      I_Contact( "HMI".LungoMacchiato )
      I_Contact( "HMI".LungoCorretto )
      I_Contact( "HMI".LungoMacchiatoCorretto )
      Move(in := 4, out1 => "Sistema".BevandaSelezionata)
   END_RUNG
   RUNG wire#w1
      I_Contact( "HMI".Corto )
      I_Contact( "HMI".CortoMacchiato )
      I_Contact( "HMI".CortoCorretto )
      I_Contact( "HMI".CortoMacchiatoCorretto )
      P_Contact(operand := "HMI".Lungo, bit := "Sistema".PLungo)
      I_Contact( "HMI".LungoMacchiato )
      I_Contact( "HMI".LungoCorretto )
      I_Contact( "HMI".LungoMacchiatoCorretto )
      Move(in := 5, out1 => "Sistema".BevandaSelezionata)
   END_RUNG
   RUNG wire#w1
      I_Contact( "HMI".Corto )
      I_Contact( "HMI".CortoMacchiato )
      I_Contact( "HMI".CortoCorretto )
      I_Contact( "HMI".CortoMacchiatoCorretto )
      I_Contact( "HMI".Lungo )
      P_Contact(operand := "HMI".LungoMacchiato, bit := "Sistema".PLungoMacchiato)
      I_Contact( "HMI".LungoCorretto )
      I_Contact( "HMI".LungoMacchiatoCorretto )
      Move(in := 6, out1 => "Sistema".BevandaSelezionata)
   END_RUNG
   RUNG wire#w1
      I_Contact( "HMI".Corto )
      I_Contact( "HMI".CortoMacchiato )
      I_Contact( "HMI".CortoCorretto )
      I_Contact( "HMI".CortoMacchiatoCorretto )
      I_Contact( "HMI".Lungo )
      I_Contact( "HMI".LungoMacchiato )
      P_Contact(operand := "HMI".LungoCorretto, bit := "Sistema".PLungoCorretto)
      I_Contact( "HMI".LungoMacchiatoCorretto )
      Move(in := 7, out1 => "Sistema".BevandaSelezionata)
   END_RUNG
   RUNG wire#w1
      I_Contact( "HMI".Corto )
      I_Contact( "HMI".CortoMacchiato )
      I_Contact( "HMI".CortoCorretto )
      I_Contact( "HMI".CortoMacchiatoCorretto )
      I_Contact( "HMI".Lungo )
      I_Contact( "HMI".LungoMacchiato )
      I_Contact( "HMI".LungoCorretto )
      P_Contact(operand := "HMI".LungoMacchiatoCorretto, bit := "Sistema".PLungoMacchiatoCorretto)
      Move(in := 8, out1 => "Sistema".BevandaSelezionata)
   END_RUNG
   RUNG wire#w1
      "ValutazioneInsufficienzaCredito"(BevandaSelezionata := "Sistema".BevandaSelezionata, CreditoUtente := "HMI".Credito, CreditoInsufficiente := "HMI".CreditoInsufficiente)
   END_RUNG
   // the same network as SCL:
   #_w1 := NOT "Sistema".BloccoInterfacciaUtente;
   #_w2 := #_w1 AND "HMI".Corto AND NOT "Sistema".PCorto;   // rising edge of "HMI".Corto
   "Sistema".PCorto := "HMI".Corto;
   IF #_w2 AND NOT "HMI".CortoMacchiato AND NOT "HMI".CortoCorretto AND NOT "HMI".CortoMacchiatoCorretto AND NOT "HMI".Lungo AND NOT "HMI".LungoMacchiato AND NOT "HMI".LungoCorretto AND NOT "HMI".LungoMacchiatoCorretto THEN
       "Sistema".BevandaSelezionata := 1;
   END_IF;
   #_w3 := #_w1 AND NOT "HMI".Corto AND "HMI".CortoMacchiato AND NOT "Sistema".PCortoMacchiato;   // rising edge of "HMI".CortoMacchiato
   "Sistema".PCortoMacchiato := "HMI".CortoMacchiato;
   IF #_w3 AND NOT "HMI".CortoCorretto AND NOT "HMI".CortoMacchiatoCorretto AND NOT "HMI".Lungo AND NOT "HMI".LungoMacchiato AND NOT "HMI".LungoCorretto AND NOT "HMI".LungoMacchiatoCorretto THEN
       "Sistema".BevandaSelezionata := 2;
   END_IF;
   #_w4 := #_w1 AND NOT "HMI".Corto AND NOT "HMI".CortoMacchiato AND "HMI".CortoCorretto AND NOT "Sistema".PCortoCorretto;   // rising edge of "HMI".CortoCorretto
   "Sistema".PCortoCorretto := "HMI".CortoCorretto;
   IF #_w4 AND NOT "HMI".CortoMacchiatoCorretto AND NOT "HMI".Lungo AND NOT "HMI".LungoMacchiato AND NOT "HMI".LungoCorretto AND NOT "HMI".LungoMacchiatoCorretto THEN
       "Sistema".BevandaSelezionata := 3;
   END_IF;
   #_w5 := #_w1 AND NOT "HMI".Corto AND NOT "HMI".CortoMacchiato AND NOT "HMI".CortoCorretto AND "HMI".CortoMacchiatoCorretto AND NOT "Sistema".PCortoMacchiatoCorretto;   // rising edge of "HMI".CortoMacchiatoCorretto
   "Sistema".PCortoMacchiatoCorretto := "HMI".CortoMacchiatoCorretto;
   IF #_w5 AND NOT "HMI".Lungo AND NOT "HMI".LungoMacchiato AND NOT "HMI".LungoCorretto AND NOT "HMI".LungoMacchiatoCorretto THEN
       "Sistema".BevandaSelezionata := 4;
   END_IF;
   #_w6 := #_w1 AND NOT "HMI".Corto AND NOT "HMI".CortoMacchiato AND NOT "HMI".CortoCorretto AND NOT "HMI".CortoMacchiatoCorretto AND "HMI".Lungo AND NOT "Sistema".PLungo;   // rising edge of "HMI".Lungo
   "Sistema".PLungo := "HMI".Lungo;
   IF #_w6 AND NOT "HMI".LungoMacchiato AND NOT "HMI".LungoCorretto AND NOT "HMI".LungoMacchiatoCorretto THEN
       "Sistema".BevandaSelezionata := 5;
   END_IF;
   #_w7 := #_w1 AND NOT "HMI".Corto AND NOT "HMI".CortoMacchiato AND NOT "HMI".CortoCorretto AND NOT "HMI".CortoMacchiatoCorretto AND NOT "HMI".Lungo AND "HMI".LungoMacchiato AND NOT "Sistema".PLungoMacchiato;   // rising edge of "HMI".LungoMacchiato
   "Sistema".PLungoMacchiato := "HMI".LungoMacchiato;
   IF #_w7 AND NOT "HMI".LungoCorretto AND NOT "HMI".LungoMacchiatoCorretto THEN
       "Sistema".BevandaSelezionata := 6;
   END_IF;
   #_w8 := #_w1 AND NOT "HMI".Corto AND NOT "HMI".CortoMacchiato AND NOT "HMI".CortoCorretto AND NOT "HMI".CortoMacchiatoCorretto AND NOT "HMI".Lungo AND NOT "HMI".LungoMacchiato AND "HMI".LungoCorretto AND NOT "Sistema".PLungoCorretto;   // rising edge of "HMI".LungoCorretto
   "Sistema".PLungoCorretto := "HMI".LungoCorretto;
   IF #_w8 AND NOT "HMI".LungoMacchiatoCorretto THEN "Sistema".BevandaSelezionata := 7; END_IF;
   #_w9 := #_w1 AND NOT "HMI".Corto AND NOT "HMI".CortoMacchiato AND NOT "HMI".CortoCorretto AND NOT "HMI".CortoMacchiatoCorretto AND NOT "HMI".Lungo AND NOT "HMI".LungoMacchiato AND NOT "HMI".LungoCorretto AND "HMI".LungoMacchiatoCorretto AND NOT "Sistema".PLungoMacchiatoCorretto;   // rising edge of "HMI".LungoMacchiatoCorretto
   "Sistema".PLungoMacchiatoCorretto := "HMI".LungoMacchiatoCorretto;
   IF #_w9 THEN "Sistema".BevandaSelezionata := 8; END_IF;
   IF #_w1 THEN
       "ValutazioneInsufficienzaCredito"(BevandaSelezionata := "Sistema".BevandaSelezionata,
                               CreditoUtente := "HMI".Credito,
                               CreditoInsufficiente := "HMI".CreditoInsufficiente);
   END_IF;
END_REGION

REGION Network 3
   // Regolazione zucchero
   // 
   // Min = 0 unità
   // Max = 5 unità
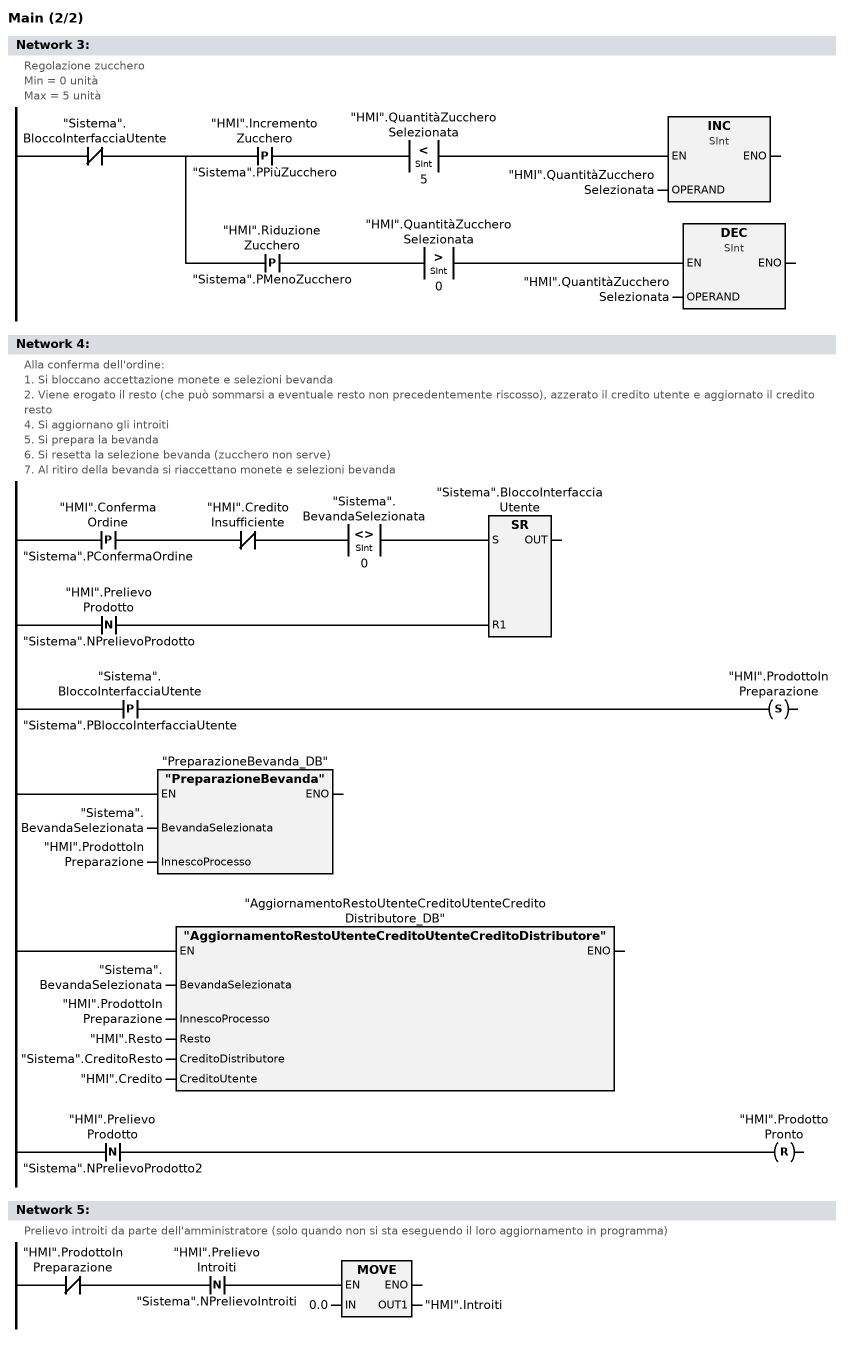
   RUNG wire#powerrail
      I_Contact( "Sistema".BloccoInterfacciaUtente )
      wire#w1
      P_Contact(operand := "HMI".IncrementoZucchero, bit := "Sistema".PPiùZucchero)
      { S7_Templates := "SrcType := SInt" } LT_Contact(in1 := "HMI".QuantitàZuccheroSelezionata, in2 := 5)
      { S7_Templates := "DestType := SInt" } Inc( "HMI".QuantitàZuccheroSelezionata )
   END_RUNG
   RUNG wire#w1
      P_Contact(operand := "HMI".RiduzioneZucchero, bit := "Sistema".PMenoZucchero)
      { S7_Templates := "SrcType := SInt" } GT_Contact(in1 := "HMI".QuantitàZuccheroSelezionata, in2 := 0)
      { S7_Templates := "DestType := SInt" } Dec( "HMI".QuantitàZuccheroSelezionata )
   END_RUNG
   // the same network as SCL:
   #_w1 := NOT "Sistema".BloccoInterfacciaUtente;
   #_w2 := #_w1 AND "HMI".IncrementoZucchero AND NOT "Sistema".PPiùZucchero;   // rising edge of "HMI".IncrementoZucchero
   "Sistema".PPiùZucchero := "HMI".IncrementoZucchero;
   IF #_w2 AND ("HMI".QuantitàZuccheroSelezionata < 5) THEN
       "HMI".QuantitàZuccheroSelezionata := "HMI".QuantitàZuccheroSelezionata + 1;
   END_IF;
   #_w3 := #_w1 AND "HMI".RiduzioneZucchero AND NOT "Sistema".PMenoZucchero;   // rising edge of "HMI".RiduzioneZucchero
   "Sistema".PMenoZucchero := "HMI".RiduzioneZucchero;
   IF #_w3 AND ("HMI".QuantitàZuccheroSelezionata > 0) THEN
       "HMI".QuantitàZuccheroSelezionata := "HMI".QuantitàZuccheroSelezionata - 1;
   END_IF;
END_REGION

REGION Network 4
   // Alla conferma dell'ordine:
   // 
   // 1. Si bloccano accettazione monete e selezioni bevanda
   // 2. Viene erogato il resto (che può sommarsi a eventuale resto non precedentemente riscosso), azzerato il credito utente e aggiornato il credito resto
   // 4. Si aggiornano gli introiti
   // 5. Si prepara la bevanda
   // 6. Si resetta la selezione bevanda (zucchero non serve)
   // 7. Al ritiro della bevanda si riaccettano monete e selezioni bevanda
   RUNG wire#powerrail
      P_Contact(operand := "HMI".ConfermaOrdine, bit := "Sistema".PConfermaOrdine)
      I_Contact( "HMI".CreditoInsufficiente )
      { S7_Templates := "SrcType := SInt" } NE_Contact(in1 := "Sistema".BevandaSelezionata, in2 := 0)
      S_SR(operand := "Sistema".BloccoInterfacciaUtente, r1 := wire#w1)
   END_RUNG
   RUNG wire#powerrail
      N_Contact(operand := "HMI".PrelievoProdotto, bit := "Sistema".NPrelievoProdotto)
   END_RUNG wire#w1
   RUNG wire#powerrail
      P_Contact(operand := "Sistema".BloccoInterfacciaUtente, bit := "Sistema".PBloccoInterfacciaUtente)
      S_Coil( "HMI".ProdottoInPreparazione )
   END_RUNG
   RUNG wire#powerrail
      "PreparazioneBevanda_DB"(BevandaSelezionata := "Sistema".BevandaSelezionata, InnescoProcesso := "HMI".ProdottoInPreparazione)
   END_RUNG
   RUNG wire#powerrail
      "AggiornamentoRestoUtenteCreditoUtenteCreditoDistributore_DB"(BevandaSelezionata := "Sistema".BevandaSelezionata, InnescoProcesso := "HMI".ProdottoInPreparazione, Resto := "HMI".Resto, CreditoDistributore := "Sistema".CreditoResto, CreditoUtente := "HMI".Credito)
   END_RUNG
   RUNG wire#powerrail
      N_Contact(operand := "HMI".PrelievoProdotto, bit := "Sistema".NPrelievoProdotto2)
      R_Coil( "HMI".ProdottoPronto )
   END_RUNG
   // the same network as SCL:
   #_w1 := "HMI".ConfermaOrdine AND NOT "Sistema".PConfermaOrdine;   // rising edge of "HMI".ConfermaOrdine
   "Sistema".PConfermaOrdine := "HMI".ConfermaOrdine;
   #_w2 := NOT "HMI".PrelievoProdotto AND "Sistema".NPrelievoProdotto;   // falling edge of "HMI".PrelievoProdotto
   "Sistema".NPrelievoProdotto := "HMI".PrelievoProdotto;
   IF #_w1 AND NOT "HMI".CreditoInsufficiente AND ("Sistema".BevandaSelezionata <> 0) THEN
       "Sistema".BloccoInterfacciaUtente := TRUE;   // SR flip-flop
   END_IF;
   IF #_w2 THEN "Sistema".BloccoInterfacciaUtente := FALSE; END_IF;
   #_w3 := "Sistema".BloccoInterfacciaUtente AND NOT "Sistema".PBloccoInterfacciaUtente;   // rising edge of "Sistema".BloccoInterfacciaUtente
   "Sistema".PBloccoInterfacciaUtente := "Sistema".BloccoInterfacciaUtente;
   IF #_w3 THEN "HMI".ProdottoInPreparazione := TRUE; END_IF;
   "PreparazioneBevanda_DB"(BevandaSelezionata := "Sistema".BevandaSelezionata,   // "PreparazioneBevanda"
                           InnescoProcesso := "HMI".ProdottoInPreparazione);
   "AggiornamentoRestoUtenteCreditoUtenteCreditoDistributore_DB"(BevandaSelezionata := "Sistema".BevandaSelezionata,   // "AggiornamentoRestoUtenteCreditoUtenteCreditoDistributore"
                           InnescoProcesso := "HMI".ProdottoInPreparazione,
                           Resto := "HMI".Resto,
                           CreditoDistributore := "Sistema".CreditoResto,
                           CreditoUtente := "HMI".Credito);
   #_w4 := NOT "HMI".PrelievoProdotto AND "Sistema".NPrelievoProdotto2;   // falling edge of "HMI".PrelievoProdotto
   "Sistema".NPrelievoProdotto2 := "HMI".PrelievoProdotto;
   IF #_w4 THEN "HMI".ProdottoPronto := FALSE; END_IF;
END_REGION

REGION Network 5
   // Prelievo introiti da parte dell'amministratore (solo quando non si sta eseguendo il loro aggiornamento in programma)
   RUNG wire#powerrail
      I_Contact( "HMI".ProdottoInPreparazione )
      N_Contact(operand := "HMI".PrelievoIntroiti, bit := "Sistema".NPrelievoIntroiti)
      Move(in := 0.0, out1 => "HMI".Introiti)
   END_RUNG
   // the same network as SCL:
   #_w1 := NOT "HMI".ProdottoInPreparazione AND NOT "HMI".PrelievoIntroiti AND "Sistema".NPrelievoIntroiti;   // falling edge of "HMI".PrelievoIntroiti
   "Sistema".NPrelievoIntroiti := "HMI".PrelievoIntroiti;
   IF #_w1 THEN "HMI".Introiti := 0.0; END_IF;
END_REGION
END_ORGANIZATION_BLOCK

(* ===== HMI "HMI_RT_1" =====
system functions are stored by id; their names below are inferred from use
connection "HMI_Collegamento_1": ETHERNET, SMART_S7_1200_OMS

HMI tags "Tabella delle variabili standard"
   "Variabile_Numero di pagina" : UInt, internal
   "HMI_ProdottoPronto" : Bool = PLC HMI.ProdottoPronto, 100 ms
   "HMI_PrelievoProdotto" : Bool = PLC HMI.PrelievoProdotto, 100 ms
   "HMI_BicchieriScarico" : Bool = PLC HMI.BicchieriScarico, 100 ms
   "HMI_PaletteScarico" : Bool = PLC HMI.PaletteScarico, 100 ms
   "HMI_CaffèScarico" : Bool = PLC HMI.CaffèScarico, 100 ms
   "HMI_LatteScarico" : Bool = PLC HMI.LatteScarico, 100 ms
   "HMI_GrappaScarico" : Bool = PLC HMI.GrappaScarico, 100 ms
   "HMI_ZuccheroScarico" : Bool = PLC HMI.ZuccheroScarico, 100 ms
   "HMI_Bicchieri" : Int = PLC HMI.Bicchieri, 100 ms
   "HMI_Palette" : Int = PLC HMI.Palette, 100 ms
   "HMI_Caffè" : SInt = PLC HMI.Caffè, 100 ms
   "HMI_Latte" : SInt = PLC HMI.Latte, 100 ms
   "HMI_Grappa" : SInt = PLC HMI.Grappa, 100 ms
   "HMI_Zucchero" : SInt = PLC HMI.Zucchero, 100 ms
   "HMI_Credito" : Real = PLC HMI.Credito, 100 ms
   "HMI_Introiti" : Real = PLC HMI.Introiti, 100 ms
   "HMI_PrelievoIntroiti" : Bool = PLC HMI.PrelievoIntroiti, 100 ms
   "HMI_CreditoInsufficiente" : Bool = PLC HMI.CreditoInsufficiente, 100 ms
   "HMI_I5cents" : Bool = PLC HMI.I5cents, 100 ms
   "HMI_I10Cents" : Bool = PLC HMI.I10Cents, 100 ms
   "HMI_I20Cents" : Bool = PLC HMI.I20Cents, 100 ms
   "HMI_I50Cents" : Bool = PLC HMI.I50Cents, 100 ms
   "HMI_I1Euro" : Bool = PLC HMI.I1Euro, 100 ms
   "HMI_I2Euro" : Bool = PLC HMI.I2Euro, 100 ms
   "HMI_Corto" : Bool = PLC HMI.Corto, 100 ms
   "HMI_CortoMacchiato" : Bool = PLC HMI.CortoMacchiato, 100 ms
   "HMI_CortoCorretto" : Bool = PLC HMI.CortoCorretto, 100 ms
   "HMI_CortoMacchiatoCorretto" : Bool = PLC HMI.CortoMacchiatoCorretto, 100 ms
   "HMI_Lungo" : Bool = PLC HMI.Lungo, 100 ms
   "HMI_LungoMacchiato" : Bool = PLC HMI.LungoMacchiato, 100 ms
   "HMI_LungoCorretto" : Bool = PLC HMI.LungoCorretto, 100 ms
   "HMI_LungoMacchiatoCorretto" : Bool = PLC HMI.LungoMacchiatoCorretto, 100 ms
   "HMI_ValvolaBicchiere" : Bool = PLC HMI.ValvolaBicchiere, 100 ms
   "HMI_ValvolaZucchero" : Bool = PLC HMI.ValvolaZucchero, 100 ms
   "HMI_ValvolaGrappa" : Bool = PLC HMI.ValvolaGrappa, 100 ms
   "HMI_ValvolaLatte" : Bool = PLC HMI.ValvolaLatte, 100 ms
   "HMI_ValvolaCaffè" : Bool = PLC HMI.ValvolaCaffè, 100 ms
   "HMI_ValvolaPaletta" : Bool = PLC HMI.ValvolaPaletta, 100 ms
   "HMI_QuantitàZuccheroSelezionata" : SInt = PLC HMI.QuantitàZuccheroSelezionata, 100 ms
   "HMI_RiduzioneZucchero" : Bool = PLC HMI.RiduzioneZucchero, 100 ms
   "HMI_IncrementoZucchero" : Bool = PLC HMI.IncrementoZucchero, 100 ms
   "HMI_ConfermaOrdine" : Bool = PLC HMI.ConfermaOrdine, 100 ms
   "HMI_Resto" : RestoUtente = PLC HMI.Resto, 100 ms
   "HMI_Resto_5Cents" : SInt = PLC HMI.Resto.5Cents, 100 ms
   "HMI_Resto_10Cents" : SInt = PLC HMI.Resto.10Cents, 100 ms
   "HMI_Resto_20Cents" : SInt = PLC HMI.Resto.20Cents, 100 ms
   "HMI_Resto_50Cents" : SInt = PLC HMI.Resto.50Cents, 100 ms
   "HMI_Resto_1Euro" : SInt = PLC HMI.Resto.1Euro, 100 ms
   "HMI_Resto_2Euro" : SInt = PLC HMI.Resto.2Euro, 100 ms
   "HMI_ProdottoInPreparazione" : Bool = PLC HMI.ProdottoInPreparazione, 100 ms

text list "Elenco testi_Nome della pagina": 1 'Pagina base'; 2 'Gestione utenti'

Template "Modello_1" 800x480
   Button "Pagina iniziale" at 1,39 size 55x39; TextOff 'Pagina iniziale'; PictureOff "NavigateHome_KTP900_Basic_PN_TR"; PictureOn "NavigateHome_KTP900_Basic_PN_TR"
      on Release: ActivateScreen("Distributore", 0)
   Button "Template_Button" at 1,79 size 55x39; TextOff 'Text'
   Button "Template_Button_1" at 1,119 size 55x39; TextOff 'Text'
   Button "Template_Button_2" at 1,159 size 55x39; TextOff 'Text'
   Button "Template_Button_3" at 1,199 size 55x39; TextOff 'Text'
   Button "Template_Button_4" at 1,239 size 55x39; TextOff 'Text'
   Button "Template_Button_5" at 1,279 size 55x39; TextOff 'Text'
   Button "Template_Button_6" at 1,319 size 55x39; TextOff 'Text'
   Button "Template_Button_7" at 1,359 size 55x39; TextOff 'Text'
   Button "Connessione" at 1,399 size 55x39; TextOff 'Connessione'; PictureOff "Login_KTP900_Basic_PN_TR"; PictureOn "Login_KTP900_Basic_PN_TR"
      on Release: function_a2a04561()
   Button "Esci" at 1,439 size 55x39; TextOff 'Esci'; PictureOff "ExitRuntime_KTP900_Basic_PN_TR"; PictureOn "ExitRuntime_KTP900_Basic_PN_TR"
      on Release: StopRuntime(0)
   SymbolicIOField "Pagina_campo_IO_simbolico" at 2,7 size 691x26; TextOff '0'; TextOn '1'; TextList "Elenco testi_Nome della pagina"
      ProcessValue <- "Variabile_Numero di pagina"
      on Change: ActivateScreenByNumber("Variabile_Numero di pagina", 0)
   DateTimeField "HmiScreenItemData" at 695,20 size 105x20
   DateTimeField "HmiScreenItemData_1" at 695,0 size 105x20

screen "Distributore" 800x480, template "Modello_1"
   on GenerateScreen: SetTag("Variabile_Numero di pagina", 1)
   Button "Pulsante_1" at 77,61 size 96x32; TextOff '0,05€'; TextOn '0,05'
      on Press: SetBit("HMI_I5cents")
      on Release: ResetBit("HMI_I5cents")
   TextField "Casella di testo_1" at 59,39 size 133x20; Text 'Inserimento credito'
   Button "Pulsante_2" at 77,93 size 96x32; TextOff '0,10€'; TextOn '0,10'
      on Press: SetBit("HMI_I10Cents")
      on Release: ResetBit("HMI_I10Cents")
   Button "Pulsante_3" at 77,125 size 96x32; TextOff '0,20€'; TextOn '0,20'
      on Press: SetBit("HMI_I20Cents")
      on Release: ResetBit("HMI_I20Cents")
   Button "Pulsante_4" at 77,157 size 96x32; TextOff '0,50€'; TextOn '0,50'
      on Press: SetBit("HMI_I50Cents")
      on Release: ResetBit("HMI_I50Cents")
   Button "Pulsante_5" at 77,189 size 96x32; TextOff '1€'; TextOn '1'
      on Press: SetBit("HMI_I1Euro")
      on Release: ResetBit("HMI_I1Euro")
   Button "Pulsante_6" at 77,221 size 96x32; TextOff '2€'; TextOn '2'
      on Press: SetBit("HMI_I2Euro")
      on Release: ResetBit("HMI_I2Euro")
   TextField "Casella di testo_2" at 310,41 size 96x20; Text 'Prelievo resto'
   Button "Pulsante_7" at 292,66 size 60x60; TextOff 'Text'; PictureOff "5cents"; PictureOn "5cents"
      on Click: function_b9b71300("HMI_Resto_5Cents", 1)
      Visibility <- "HMI_Resto_5Cents"
   Button "Pulsante_8" at 368,66 size 60x60; TextOff 'Text'; PictureOff "10cents"; PictureOn "10cents"
      on Click: function_b9b71300("HMI_Resto_10Cents", 1)
      Visibility <- "HMI_Resto_10Cents"
   Button "Pulsante_9" at 292,134 size 60x60; TextOff 'Text'; PictureOff "20cents"; PictureOn "20cents"
      on Click: function_b9b71300("HMI_Resto_20Cents", 1)
      Visibility <- "HMI_Resto_20Cents"
   Button "Pulsante_10" at 368,134 size 60x60; TextOff 'Text'; PictureOff "50cents"; PictureOn "50cents"
      on Click: function_b9b71300("HMI_Resto_50Cents", 1)
      Visibility <- "HMI_Resto_50Cents"
   Button "Pulsante_11" at 292,204 size 60x60; TextOff 'Text'; PictureOff "1euro"; PictureOn "1euro"
      on Click: function_b9b71300("HMI_Resto_1Euro", 1)
      Visibility <- "HMI_Resto_1Euro"
   Button "Pulsante_12" at 368,204 size 60x60; TextOff 'Text'; PictureOff "2euro"; PictureOn "2euro"
      on Click: function_b9b71300("HMI_Resto_2Euro", 1)
      Visibility <- "HMI_Resto_2Euro"
   IOField "Campo I/O_1" at 245,83 size 37x32; FormatPattern 99
      ProcessValue <- "HMI_Resto_5Cents"
   IOField "Campo I/O_2" at 245,147 size 37x32; FormatPattern 99
      ProcessValue <- "HMI_Resto_20Cents"
   IOField "Campo I/O_3" at 245,216 size 37x32; FormatPattern 99
      ProcessValue <- "HMI_Resto_1Euro"
   IOField "Campo I/O_4" at 440,83 size 37x32; FormatPattern 99
      ProcessValue <- "HMI_Resto_10Cents"
   IOField "Campo I/O_5" at 440,147 size 37x32; FormatPattern 99
      ProcessValue <- "HMI_Resto_50Cents"
   IOField "Campo I/O_6" at 440,216 size 37x32; FormatPattern 99
      ProcessValue <- "HMI_Resto_2Euro"
   IOField "Campo I/O_7" at 100,278 size 49x32; FormatPattern 99.99
      ProcessValue <- "HMI_Credito"
      Appearance <- "HMI_CreditoInsufficiente"
   TextField "Casella di testo_3" at 96,257 size 52x20; Text 'Credito'
   Group "Group" at 566,286 size 89x83; Picture "Grafica_6"
   Group "Group_1" at 566,174 size 89x83; Picture "Grafica_6"
   Group "Group_3" at 701,286 size 89x83; Picture "Grafica_6"
   Group "Group_4" at 701,174 size 89x83; Picture "Grafica_6"
   Group "Group_5" at 701,64 size 89x83; Picture "Grafica_6"
   TextField "Casella di testo_5" at 701,43 size 52x20; Text 'Paletta'
   TextField "Casella di testo_6" at 572,152 size 39x20; Text 'Caffè'
   TextField "Casella di testo_7" at 707,154 size 40x20; Text 'Latte'
   TextField "Casella di testo_8" at 566,266 size 51x20; Text 'Grappa'
   TextField "Casella di testo_9" at 695,266 size 64x20; Text 'Zucchero'
   Group "Group_6" at 562,44 size 93x103; Picture "Grafica_6"
   Button "Pulsante_13" at 617,372 size 82x82; TextOff 'Text'; PictureOff "BevandaPronta"; PictureOn "BevandaPronta_1"
      Visibility <- "HMI_ProdottoPronto"
      on Press: SetBit("HMI_PrelievoProdotto")
      on Release: ResetBit("HMI_PrelievoProdotto")
   GraphicView "Vista grafica_19" at 588,375 size 145x76; Picture "PaoloBitta"
      Visibility <- "HMI_ProdottoInPreparazione"
   TextField "Casella di testo_10" at 322,300 size 126x20; Text 'Selezione bevanda'
   Button "Pulsante_14" at 207,323 size 175x32; TextOff 'Corto 0,30€'; TextOn 'Corto'
      on Press: SetBit("HMI_Corto")
      on Release: ResetBit("HMI_Corto")
   Button "Pulsante_15" at 382,323 size 175x32; TextOff 'Corto macchiato 0,40€'; TextOn 'Corto macchiato'
      on Press: SetBit("HMI_CortoMacchiato")
      on Release: ResetBit("HMI_CortoMacchiato")
   Button "Pulsante_16" at 382,355 size 175x32; TextOff 'Corto corretto 0,40€'; TextOn 'Corto corretto'
      on Press: SetBit("HMI_CortoCorretto")
      on Release: ResetBit("HMI_CortoCorretto")
   Button "Pulsante_17" at 207,355 size 175x32; TextOff 'Corto macchiato corretto 0,50€'; TextOn 'Corto macchiato corretto'
      on Press: SetBit("HMI_CortoMacchiatoCorretto")
      on Release: ResetBit("HMI_CortoMacchiatoCorretto")
   Button "Pulsante_18" at 207,391 size 175x32; TextOff 'Lungo 0,60€'; TextOn 'Lungo'
      on Press: SetBit("HMI_Lungo")
      on Release: ResetBit("HMI_Lungo")
   Button "Pulsante_19" at 382,391 size 175x32; TextOff 'Lungo macchiato 0,70€'; TextOn 'Lungo macchiato'
      on Release: ResetBit("HMI_LungoMacchiato")
      on Press: SetBit("HMI_LungoMacchiato")
   Button "Pulsante_20" at 382,423 size 175x32; TextOff 'Lungo corretto 0,70€'; TextOn 'Lungo corretto'
      on Press: SetBit("HMI_LungoCorretto")
      on Release: ResetBit("HMI_LungoCorretto")
   Button "Pulsante_21" at 207,423 size 175x32; TextOff 'Lungo macchiato corretto 0,80€'; TextOn 'Lungo macchiato corretto'
      on Press: SetBit("HMI_LungoMacchiatoCorretto")
      on Release: ResetBit("HMI_LungoMacchiatoCorretto")
   TextField "Casella di testo_11" at 59,328 size 146x20; Text 'Regolazione zucchero'
   Button "Pulsante_22" at 65,355 size 38x32; TextOff '-'
      on Press: SetBit("HMI_RiduzioneZucchero")
      on Release: ResetBit("HMI_RiduzioneZucchero")
   Button "Pulsante_23" at 161,355 size 37x32; TextOff '+'
      on Release: ResetBit("HMI_IncrementoZucchero")
      on Press: SetBit("HMI_IncrementoZucchero")
   IOField "Campo I/O_8" at 114,355 size 36x32; FormatPattern 9
      ProcessValue <- "HMI_QuantitàZuccheroSelezionata"
   Button "Pulsante_24" at 73,422 size 119x32; TextOff 'Conferma ordine'
      on Press: SetBit("HMI_ConfermaOrdine")
      on Release: ResetBit("HMI_ConfermaOrdine")
   Button "Button_1" at 1,360 size 54x37; TextOff 'IA'; TextOn 'InfoAdmin'; Authorization "Visualizzazione introiti"
      on Click: ActivateScreen("InfoAdmin", 0)
   GraphicView "Vista grafica_10" at 566,286 size 69x83; Picture "Grafica_6"
   GraphicView "Vista grafica_9" at 622,306 size 19x43; Picture "Grafica_5"
      Visibility <- "HMI_ValvolaGrappa"
   GraphicView "Vista grafica_8" at 608,316 size 47x23; Picture "Grafica_4"
      Visibility <- "HMI_ValvolaGrappa"
   GraphicView "Vista grafica_1" at 566,174 size 69x83; Picture "Grafica_6"
   GraphicView "Vista grafica_2" at 622,194 size 19x43; Picture "Grafica_5"
      Visibility <- "HMI_ValvolaCaffè"
   GraphicView "Vista grafica_3" at 608,204 size 47x23; Picture "Grafica_4"
      Visibility <- "HMI_ValvolaCaffè"
   GraphicView "Vista grafica_4" at 566,64 size 69x83; Picture "Grafica_6"
   GraphicView "Vista grafica_5" at 622,84 size 19x43; Picture "Grafica_5"
      Visibility <- "HMI_ValvolaBicchiere"
   GraphicView "Vista grafica_6" at 608,94 size 47x23; Picture "Grafica_4"
      Visibility <- "HMI_ValvolaBicchiere"
   Group "Group_2" at 566,64 size 89x83; Picture "Grafica_6"
   TextField "Casella di testo_4" at 562,44 size 63x20; Text 'Bicchiere'
   GraphicView "Vista grafica_7" at 701,286 size 69x83; Picture "Grafica_6"
   GraphicView "Vista grafica_11" at 757,306 size 19x43; Picture "Grafica_5"
      Visibility <- "HMI_ValvolaZucchero"
   GraphicView "Vista grafica_12" at 743,316 size 47x23; Picture "Grafica_4"
      Visibility <- "HMI_ValvolaZucchero"
   GraphicView "Vista grafica_13" at 701,174 size 69x83; Picture "Grafica_6"
   GraphicView "Vista grafica_14" at 757,194 size 19x43; Picture "Grafica_5"
      Visibility <- "HMI_ValvolaLatte"
   GraphicView "Vista grafica_15" at 743,204 size 47x23; Picture "Grafica_4"
      Visibility <- "HMI_ValvolaLatte"
   GraphicView "Vista grafica_16" at 701,64 size 69x83; Picture "Grafica_6"
   GraphicView "Vista grafica_17" at 757,84 size 19x43; Picture "Grafica_5"
      Visibility <- "HMI_ValvolaPaletta"
   GraphicView "Vista grafica_18" at 743,94 size 47x23; Picture "Grafica_4"
      Visibility <- "HMI_ValvolaPaletta"

screen "Gestione utenti" 800x480, template "Modello_1"
   on GenerateScreen: SetTag("Variabile_Numero di pagina", 2)
   UserView "HmiScreenItemData" at 57,89 size 740x383
   Button "Indietro" at 57,41 size 159x47; TextOff 'Indietro'
      on Release: ActivateScreen("Distributore", 0)

screen "Serbatoi" 800x480
   Bar "Barra grafica_1" at 647,86 size 100x200; MinimumValue 0; MaximumValue 100
      ProcessValue <- "HMI_Zucchero"
   Bar "Barra grafica_2" at 498,85 size 100x200; MinimumValue 0; MaximumValue 100
      ProcessValue <- "HMI_Grappa"
   Bar "Barra grafica_3" at 357,84 size 100x200; MinimumValue 0; MaximumValue 100
      ProcessValue <- "HMI_Latte"
   Bar "Barra grafica_4" at 234,84 size 100x200; MinimumValue 0; MaximumValue 100
      ProcessValue <- "HMI_Caffè"
   IOField "Campo I/O_1" at 90,108 size 96x32; FormatPattern 99999
      ProcessValue <- "HMI_Bicchieri"
   IOField "Campo I/O_2" at 87,200 size 96x32; FormatPattern 99999
      ProcessValue <- "HMI_Palette"
   TextField "Casella di testo_1" at 106,84 size 58x20; Text 'Bicchieri'
   TextField "Casella di testo_2" at 105,178 size 52x20; Text 'Palette'
   TextField "Casella di testo_3" at 262,58 size 39x20; Text 'Caffè'
   TextField "Casella di testo_4" at 387,58 size 40x20; Text 'Latte'
   TextField "Casella di testo_5" at 524,58 size 51x20; Text 'Grappa'
   TextField "Casella di testo_6" at 668,58 size 64x20; Text 'Zucchero'
   GraphicIOField "PlotLight_Square_N_Mono" at 21,92 size 50x50; PictureOff "PilotLight_Square_N_Off_mono"; PictureOn "PilotLight_Square_N_On_mono"
      ProcessValue <- "HMI_BicchieriScarico"
      Appearance <- "HMI_BicchieriScarico"
   GraphicIOField "PlotLight_Square_N_Mono_1" at 259,293 size 50x50; PictureOff "PilotLight_Square_N_Off_mono"; PictureOn "PilotLight_Square_N_On_mono"
      ProcessValue <- "HMI_CaffèScarico"
      Appearance <- "HMI_CaffèScarico"
   GraphicIOField "PlotLight_Square_N_Mono_2" at 387,293 size 50x50; PictureOff "PilotLight_Square_N_Off_mono"; PictureOn "PilotLight_Square_N_On_mono"
      Appearance <- "HMI_LatteScarico"
      ProcessValue <- "HMI_LatteScarico"
   GraphicIOField "PlotLight_Square_N_Mono_3" at 521,292 size 50x50; PictureOff "PilotLight_Square_N_Off_mono"; PictureOn "PilotLight_Square_N_On_mono"
      ProcessValue <- "HMI_GrappaScarico"
      Appearance <- "HMI_GrappaScarico"
   GraphicIOField "PlotLight_Square_N_Mono_4" at 675,292 size 50x50; PictureOff "PilotLight_Square_N_Off_mono"; PictureOn "PilotLight_Square_N_On_mono"
      Appearance <- "HMI_ZuccheroScarico"
      ProcessValue <- "HMI_ZuccheroScarico"
   GraphicIOField "PlotLight_Square_N_Mono_5" at 19,186 size 50x50; PictureOff "PilotLight_Square_N_Off_mono"; PictureOn "PilotLight_Square_N_On_mono"
      ProcessValue <- "HMI_PaletteScarico"
      Appearance <- "HMI_PaletteScarico"

screen "InfoAdmin" 800x480
   TextField "Casella di testo_1" at 64,27 size 50x20; Text 'Introiti'
   IOField "Campo I/O_1" at 37,52 size 108x32; FormatPattern 9.99e
      ProcessValue <- "HMI_Introiti"
   Button "Pulsante_1" at 159,52 size 96x32; TextOff 'Prelievo'; Authorization "Prelievo introiti"
      on Press: SetBit("HMI_PrelievoIntroiti")
      on Release: ResetBit("HMI_PrelievoIntroiti")
   Button "Button_1" at 37,234 size 192x32; TextOff 'Distributore'
      on Click: ActivateScreen("Distributore", 0)
*)